  # ITEM_MAP.append(create_item(id=31, ls_item="TestLM", frame=TestLM, actionlist=[ActionManipulator.PICK, ActionManipulator.PLACE], item_model=create_item_model(inner=Rack.SYSMEX_CS2500), lm_id=5, description="LM Test"))
  # Fills the Vision Config List with Projectrelated Data
  # workspaceid and skillid are highly robominds related so probably will not stay like this in the future
  # sample detection: dx and dy are used to calculate the positions in a rack and given by the offset which will be applied in order to assign the sample to a place in the rack
  # create_vision_config(workspace_id="", skill_id="", item_id=-1, capture_pos=p[0,0,0,0,0,0], dx=0, dy=0, target_origin=p[0,0,0,0,0,0], selector="default", description="default")
  # VISION_CONFIG_MAP.append(create_vision_config(workspace_id="96017791-f581-4e9e-93da-6951695fccc8", skill_id="8885cfe1-6784-4293-bd26-52ebdc67bf95", capture_pos=F10_Cap_CF, target_origin=p[0,0,0,0,0,0], item_id=11, description="LM Detect CF"))
  # VISION_CONFIG_MAP.append(create_vision_config(workspace_id="96017791-f581-4e9e-93da-6951695fccc8", skill_id="8885cfe1-6784-4293-bd26-52ebdc67bf95", capture_pos=F8_Cap_Cobas_LM, target_origin=p[0,0,0,0,0,0], item_id=8, description="LM Detect Cobas Racks"))
  # VISION_CONFIG_MAP.append(create_vision_config(workspace_id="8f0ad01c-dc36-4fdd-b295-0b6b4a38b89a", skill_id="afdc9e13-ea83-40d6-a805-bb041453d2e5", capture_pos=F3_Cap_Input, target_origin=F2_uLM_Input, item_id=3, description="Lab Solution Input Capture"))
  # VISION_CONFIG_MAP.append(create_vision_config(workspace_id="96017791-f581-4e9e-93da-6951695fccc8", skill_id="8885cfe1-6784-4293-bd26-52ebdc67bf95", capture_pos=F19_XN550_Cap, target_origin=F18_XN550_Input, item_id=18, description="Input XN550"))
  # VISION_CONFIG_MAP.append(create_vision_config(workspace_id="96017791-f581-4e9e-93da-6951695fccc8", skill_id="8885cfe1-6784-4293-bd26-52ebdc67bf95", capture_pos=F19_XN550_Cap, target_origin=POS_Z, item_id=19, description="LM Detect XN550F"))
  # VISION_CONFIG_MAP.append(create_vision_config(workspace_id="96017791-f581-4e9e-93da-6951695fccc8", skill_id="8885cfe1-6784-4293-bd26-52ebdc67bf95", capture_pos=F10_Cap_CF, target_origin=POS_Z, item_id=10, description="LM Detect CF"))
  # VISION_CONFIG_MAP.append(create_vision_config(workspace_id="96017791-f581-4e9e-93da-6951695fccc8", skill_id="8885cfe1-6784-4293-bd26-52ebdc67bf95", capture_pos=F19_XN550_Cap, target_origin=F20_XN550_Draw, item_id=20, description="Drawer XN550"))
  # VISION_CONFIG_MAP.append(create_vision_config(workspace_id="96017791-f581-4e9e-93da-6951695fccc8", skill_id="8885cfe1-6784-4293-bd26-52ebdc67bf95", capture_pos=F19_XN550_Cap, target_origin=F21_XN550_Btn, item_id=21, description="Button XN550"))
  # VISION_CONFIG_MAP.append(create_vision_config(workspace_id="96017791-f581-4e9e-93da-6951695fccc8", skill_id="8885cfe1-6784-4293-bd26-52ebdc67bf95", capture_pos=TestLMCap, target_origin=p[0,0,0,0,0,0], item_id=30, description="Button XN550"))
  # VISION_CONFIG_MAP.append(create_vision_config(workspace_id="96017791-f581-4e9e-93da-6951695fccc8", skill_id="8885cfe1-6784-4293-bd26-52ebdc67bf95", capture_pos=TestLMCap, target_origin=TestLM, item_id=31, description="Button XN550"))

  # VISION_CONFIG_MAP.append(create_vision_config(workspace_id="96017791-f581-4e9e-93da-6951695fccc8", skill_id="8885cfe1-6784-4293-bd26-52ebdc67bf95", target_origin=p[0,0,0,0,0,0], item_id=11, description="LM Detect CF"))
  # VISION_CONFIG_MAP.append(create_vision_config(workspace_id="96017791-f581-4e9e-93da-6951695fccc8", skill_id="8885cfe1-6784-4293-bd26-52ebdc67bf95", target_origin=p[0,0,0,0,0,0], item_id=8, description="LM Detect Cobas Racks"))
  # VISION_CONFIG_MAP.append(create_vision_config(workspace_id="8f0ad01c-dc36-4fdd-b295-0b6b4a38b89a", skill_id="afdc9e13-ea83-40d6-a805-bb041453d2e5", target_origin=F2_uLM_Input, item_id=3, description="Lab Solution Input Capture"))
  # VISION_CONFIG_MAP.append(create_vision_config(workspace_id="96017791-f581-4e9e-93da-6951695fccc8", skill_id="8885cfe1-6784-4293-bd26-52ebdc67bf95", target_origin=F18_XN550_Input, item_id=18, description="Input XN550"))
  # VISION_CONFIG_MAP.append(create_vision_config(workspace_id="96017791-f581-4e9e-93da-6951695fccc8", skill_id="8885cfe1-6784-4293-bd26-52ebdc67bf95", target_origin=POS_Z, item_id=19, description="LM Detect XN550F"))
  # VISION_CONFIG_MAP.append(create_vision_config(workspace_id="96017791-f581-4e9e-93da-6951695fccc8", skill_id="8885cfe1-6784-4293-bd26-52ebdc67bf95", target_origin=POS_Z, item_id=10, description="LM Detect CF"))
  # VISION_CONFIG_MAP.append(create_vision_config(workspace_id="96017791-f581-4e9e-93da-6951695fccc8", skill_id="8885cfe1-6784-4293-bd26-52ebdc67bf95", target_origin=F20_XN550_Draw, item_id=20, description="Drawer XN550"))
  # VISION_CONFIG_MAP.append(create_vision_config(workspace_id="96017791-f581-4e9e-93da-6951695fccc8", skill_id="8885cfe1-6784-4293-bd26-52ebdc67bf95", target_origin=F21_XN550_Btn, item_id=21, description="Button XN550"))
  # VISION_CONFIG_MAP.append(create_vision_config(workspace_id="96017791-f581-4e9e-93da-6951695fccc8", skill_id="8885cfe1-6784-4293-bd26-52ebdc67bf95", target_origin=p[0,0,0,0,0,0], item_id=30, description="Button XN550"))
  # VISION_CONFIG_MAP.append(create_vision_config(workspace_id="96017791-f581-4e9e-93da-6951695fccc8", skill_id="8885cfe1-6784-4293-bd26-52ebdc67bf95", target_origin=TestLM, item_id=31, description="Button XN550"))

  # local inputrack = find_pattern_by_name("INPUT")
  # INSPECT_CONFIG_MAP.append(create_inspect_config(item_id=3, dx=inputrack.pattern_width[0]/(inputrack.pattern_size[0]-1), dy=inputrack.pattern_width[1]/(inputrack.pattern_size[1]-1), rack_size=inputrack.pattern_size , description="Input Capture"))
  # # Fills the Landmark List with Projectrelated Data
  # # create_landmark(lm_id=0, marker_id=-1, marker_size=0.1, marker_type="aruco_7x7", capture_pos=p[0,0,0,0,0,0], init_frame=p[0,0,0,0,0,0], search_offset=[0,0,0], actual_frame=p[0,0,0,0,0,0], description="")
  # LANDMARK_MAP.append(create_landmark(lm_id=1, marker_id=3, marker_size=0.1, marker_type="aruco_7x7", capture_pos = F10_Cap_CF, init_frame=p[-0.617789, -0.065471, 0.07918, 0.020983, -0.012695, 1.512066], search_offset=[0.15, 0.15, 0.1], actual_frame=p[-0.617789, -0.065471, 0.07918, 0.020983, -0.012695, 1.512066], description="LM CF Lid"))
  # LANDMARK_MAP.append(create_landmark(lm_id=2, marker_id=-1, marker_size=0.0085, marker_type="aruco_4x4", capture_pos = F8_Cap_Cobas_LM, init_frame=p[0,0,0,0,0,0], search_offset=[0.15, 0.15, 0.1], actual_frame=POS_Z, description="LM Cobas Rack Detection"))
  # LANDMARK_MAP.append(create_landmark(lm_id=3, marker_id=0, marker_size=0.1, marker_type="aruco_7x7", capture_pos = F17_Cobas_Cap, init_frame=p[-0.667,-0.194,0.100,0,0,0], search_offset=[0.15, 0.15, 0.1], actual_frame=POS_Z, description="LM Cobas Cap"))
  # LANDMARK_MAP.append(create_landmark(lm_id=4, marker_id=4, marker_size=0.1, marker_type="aruco_7x7", capture_pos = F19_XN550_Cap, init_frame=p[0.124,-0.976,0.355,-0.008,0.025,3.131], search_offset=[0.15, 0.15, 0.1], actual_frame=p[0,0,0,0,0,0], description="LM XN550 Cap"))
  # LANDMARK_MAP.append(create_landmark(lm_id=5, marker_id=0, marker_size=0.1, marker_type="aruco_7x7", capture_pos = TestLMCap, init_frame=p[-0.49,-0.144,0.092,0,-0.008,0.001], search_offset=[0.15, 0.15, 0.1], actual_frame=POS_Z, description="LM Test"))
  # # Configuration of all movement related parameters
  # # create_movement(id=0, hh_approach=POS_Z, h_approach=POS_Z, approach=POS_Z, h_target=POS_Z, target=POS_Z, retract=POS_Z, h_retract=POS_Z, hh_retract=POS_Z, h_frame=POS_Z, frame=POS_Z, speed=1, acceleration=1, description="default")
  # MOVEMENT_MAP.append(create_movement(description="TestLMCap", frame=TestLMCap, actionlist=[ActionManipulator.MOVE_TO]))
  # MOVEMENT_MAP.append(create_movement(description="TestLM", frame=TestLM, actionlist=[ActionManipulator.PICK,ActionManipulator.PLACE],
  #         approach=p[0,0,0.1,0,0,0],
  #         retract=p[0,0,0.1,0,0,0]))
  # MOVEMENT_MAP.append(create_movement(description="Home - MOVE_TO", frame=F1_uLM_Home, actionlist=[ActionManipulator.MOVE_TO]))
  # MOVEMENT_MAP.append(create_movement(description="Input - PICK&PLACE", frame=F2_uLM_Input, actionlist=[ActionManipulator.PICK,ActionManipulator.PLACE],
  #         approach=p[0,0,0.1,0,0,0],
  #         retract=p[0,0,0.1,0,0,0]))
  # MOVEMENT_MAP.append(create_movement(description="Capture Input - MOVE_TO", frame=F3_Cap_Input, actionlist=[ActionManipulator.MOVE_TO]))
  # MOVEMENT_MAP.append(create_movement(description="BIN - PLACE", frame=F4_uLM_Bin, actionlist=[ActionManipulator.PLACE],
  #         approach=p[0,0,0.1,0,0,0],
  #         retract=p[0,0,0.1,0,0,0]))
  # MOVEMENT_MAP.append(create_movement(description="Gripper - Move To", frame=F5_uLM_Gripper, actionlist=[ActionManipulator.MOVE_TO],
  #         approach=p[0,0,0.1,0,0,0]))
  # MOVEMENT_MAP.append(create_movement(description="Gripper - Pick", frame=F5_uLM_Gripper, actionlist=[ActionManipulator.PICK],
  #         retract=p[0,0,0.1,0,0,0]))
  # MOVEMENT_MAP.append(create_movement(description="Gripper - Place", frame=F5_uLM_Gripper, actionlist=[ActionManipulator.PLACE],
  #         approach=p[0,0,0.1,0,0,0]))
  # MOVEMENT_MAP.append(create_movement(description="CobasRack Pick & Place", frame=F6_uLM_Cobas_R, actionlist=[ActionManipulator.PICK,ActionManipulator.PLACE],
  #         approach=p[0,0,0.1,0,0,0],
  #         target=p[0,0,0,0,0,d2r(90)],
  #         retract=p[0,0,0.1,0,0,0]))
  # MOVEMENT_MAP.append(create_movement(description="CobasMagazine Pick & Place", frame=F7_uLM_Coba_Mag, actionlist=[ActionManipulator.PICK,ActionManipulator.PLACE],
  #         approach=p[0,0,0.1,0,0,0],
  #         target=p[0,0,0,0,0,-d2r(90)],
  #         retract=p[0,0,0.1,0,0,0]))
  # MOVEMENT_MAP.append(create_movement(description="Capture Position Cobas Landmarks", frame=F8_Cap_Cobas_LM, actionlist=[ActionManipulator.MOVE_TO]))
  # MOVEMENT_MAP.append(create_movement(description="TaraMagazine - PICK & PLACE", frame=F9_uLM_Tara, actionlist=[ActionManipulator.PICK,ActionManipulator.PLACE],
  #         approach=p[0,0,0.13,0,0,0],
  #         target=p[0,0,0,0,0,-d2r(90)],
  #         retract=p[0,0,0.13,0,0,0]))
  # MOVEMENT_MAP.append(create_movement(description="Capture Position - Centrifuge LM", frame=F10_Cap_CF,actionlist=[ActionManipulator.MOVE_TO]))
  # MOVEMENT_MAP.append(create_movement(description="Pick and Place Racks - Centrifuge Lid", frame=F11_CF_PiPl, actionlist=[ActionManipulator.PICK,ActionManipulator.PLACE],
  #         approach=p[0,0,0.3,0,0,0],
  #         retract=p[0,0,0.3,0,0,0]))
  # MOVEMENT_MAP.append(create_movement(description="Pick and Place Samples - Centrifuge on uLM", frame=F12_uLM_CF_Mag, actionlist=[ActionManipulator.PICK,ActionManipulator.PLACE],
  #         approach=p[0,0,0.13,0,0,0],
  #         retract=p[0,0,0.13,0,0,0]
  #         ))
  # MOVEMENT_MAP.append(create_movement(description="Pick and Place Racks - Centrifuge on uLM", frame=F13_uLM_CF_R, actionlist=[ActionManipulator.PICK,ActionManipulator.PLACE],
  #         approach=p[0,0,0.15,0,0,0],
  #         retract=p[0,0,0.15,0,0,0]
  #         ))

  # MOVEMENT_MAP.append(create_movement(description="Pick and Place Samples XN550 Racks in Device", frame=F18_XN550_Input, actionlist=[ActionManipulator.PICK,ActionManipulator.PLACE],
  #         approach=p[0,0,0.1,0,0,0],
  #         target = p[0,0,0,0,0,d2r(90)],
  #         retract=p[0,0,0.1,0,0,0]
  #         ))
  # MOVEMENT_MAP.append(create_movement(description="Capture LM XN550", frame=F19_XN550_Cap, actionlist=[ActionManipulator.MOVE_TO]))
  # MOVEMENT_MAP.append(create_movement(description="Open XN550 Drawer ", frame=F20_XN550_Draw, actionlist=[ActionManipulator.DRAWER_OPEN],
  #         h_approach=p[0.07,0,0.1,0,0,0],
  #         approach=p[0,0,0.1,0,0,0],
  #         target = p[0,0,0,0,0,d2r(90)],
  #         retract=p[0.07,0,0,0,0,0],
  #         h_retract=p[0.07,0,0.1,0,0,0]
  #         ))
  # MOVEMENT_MAP.append(create_movement(description="Close XN550 Drawer ", frame=F20_XN550_Draw, actionlist=[ActionManipulator.DRAWER_CLOSE],
  #         h_approach=p[0.07,0,0.1,0,0,0],
  #         approach=p[0.07,0,0,0,0,0],
  #         target = p[0,0,0,0,0,d2r(90)],
  #         retract=p[0,0,0.1,0,0,0],
  #         h_retract=p[0.07,0,0.1,0,0,0]
  #         ))
  # MOVEMENT_MAP.append(create_movement(description="Push XN550 Button ", frame=F21_XN550_Btn, actionlist=[ActionManipulator.PUSH],
  #         approach=p[0,0,0.15,0,0,0],
  #         retract=p[0,0,0.15,0,0,0]
  #         ))
  # MOVEMENT_MAP.append(create_movement(description="Capture Position 2 Input", frame=F_Cap_Input2,actionlist=[ActionManipulator.MOVE_TO]))



  $ 19 "Script: SCRIPT Objects V0.1.script"
  #*****************************************************
  # customer          :   INTERNAL
  # project name      :
  #****************************************************
  # controller        :   UR
  # software          :   5.17.3
  #****************************************************
  # author            :   P. Koehnke
  # Copyright (c)     :   United Robotics Group
  #                       An der Riede 2
  #                       28816 Stuhr
  #                       Germany
  #****************************************************
  # description       :   object database
  # version:      	:   0.1
  # created           :   09.10.2024
  # updated           :
  #****************************************************
  # modifications     :
  #
  # date              :
  # name              :
  # reason            :
  #****************************************************

  def create_object_2(id=0, name="", type=0, dimension=struct(length=0, width=0, height=0, diameter=0), gripper_offset=p[0,0,0,0,0,0]):
      return struct(id=id, name=name, type=type, dimension=dimension, gripper_offset=gripper_offset)
  end

  OBJ = create_object_2()
  OBJs = make_list(0, create_object_2(), 50)

  OBJs.append(create_object_2(id=1, name="rack centrifuge", type=1, dimension=struct(length=0, width=0, height=0.106, diameter=0.020), gripper_offset=p[0,0,0.095,0,0,2.356]))
  OBJs.append(create_object_2(id=2, name="sample tube 1", type=2, dimension=struct(length=0, width=0, height=0.106, diameter=0.015), gripper_offset=p[0,0,0,0,0,0]))
  OBJs.append(create_object_2(id=3, name="rack sarstedt", type=3, dimension=struct(length=0, width=0, height=0.100, diameter=0.020), gripper_offset=p[0,0,0,0,0,0]))
  OBJs.append(create_object_2(id=4, name="Lab bottle", type=4, dimension=struct(length=0, width=0, height=0.100, diameter=0.030), gripper_offset=p[0,0,0.2,0,0,0]))
  OBJs.append(create_object_2(id=5, name="Vial", type=5, dimension=struct(length=0, width=0, height=0.100, diameter=0.0275), gripper_offset=p[0,0,0,0,0,0]))
  OBJs.append(create_object_2(id=6, name="Container", type=6, dimension=struct(length=0.0, width=0.0, height=0, diameter=0.0), gripper_offset=p[0,0,0,0,0,0]))
  OBJs.append(create_object_2(id=7, name="Target_container", type=7, dimension=struct(length=0.06, width=0.06, height=0.134, diameter=0.05), gripper_offset=p[0,0,0,0,0,0]))
  OBJs.append(create_object_2(id=8, name="Spatula", type=8, dimension=struct(length=0.03, width=0.03, height=0.23, diameter=0.05), gripper_offset=p[0,0,0,0,0,0]))
  OBJs.append(create_object_2(id=9, name="rack pipet", type=9, dimension=struct(length=0.03, width=0.03, height=0.23, diameter=0.05), gripper_offset=p[0,0,0,0,0,0]))

  def create_jig_2(id=0, name="", type=0, capacity=0, jig_offset=p[0,0,0,0,0,0]):
      # iformation about used jigs
      return struct(id=id, name=name, type=type, capacity=capacity, jig_offset=jig_offset)
  end

  JIG2 = create_jig_2()
  JIGs = make_list(0, create_jig_2(), 20)

  JIGs.append(create_jig_2(id=1, name="3FG", type=1, capacity=1, jig_offset=p[0,0,0,0,0,0]))
  JIGs.append(create_jig_2(id=2, name="jig input", type=2, capacity=1, jig_offset=p[0,0,0,0,0,-3.927]))
  JIGs.append(create_jig_2(id=3, name="jig output", type=3, capacity=1, jig_offset=p[0,0,0,0,0,0.78]))
  JIGs.append(create_jig_2(id=6, name="jig bin", type=6, capacity=1, jig_offset=p[0,0,0,0,0,0]))
  JIGs.append(create_jig_2(id=7, name="jig sarstedt racks", type=7, capacity=1, jig_offset=p[0,0,-0.02,0,0,0]))
  JIGs.append(create_jig_2(id=8, name="NoK Bin", type=8, capacity=1, jig_offset=p[0,0,0,0,0,0]))
  JIGs.append(create_jig_2(id=9, name="Pick bott jig", type=9, capacity=1, jig_offset=p[0,0,0,0,0,0]))
  JIGs.append(create_jig_2(id=10, name="Place bott jig", type=10, capacity=1, jig_offset=p[0,0,0,0,0,0]))
  JIGs.append(create_jig_2(id=11, name="bottle shake jig", type=11, capacity=1, jig_offset=p[0,0,0,0,0,0]))
  JIGs.append(create_jig_2(id=12, name="Pick Vial jig", type=12, capacity=1, jig_offset=p[0,0,0,0,0,0]))
  JIGs.append(create_jig_2(id=13, name="Place Vial jig", type=13, capacity=1, jig_offset=p[0,0,0,0,0,0]))
  JIGs.append(create_jig_2(id=14, name="Liquid transfer jig", type=14, capacity=1, jig_offset=p[0,0,0,0,0,0]))
  JIGs.append(create_jig_2(id=15, name="Pick station jig", type=15, capacity=1, jig_offset=p[0,0,0,0,0,0]))
  JIGs.append(create_jig_2(id=16, name="Place station jig", type=16, capacity=1, jig_offset=p[0,0,0,0,0,0]))
  JIGs.append(create_jig_2(id=17, name="Weigh station jig", type=17, capacity=1, jig_offset=p[0,0,0,0,0,0]))
  JIGs.append(create_jig_2(id=18, name="Pick station 1", type=18, capacity=1, jig_offset=p[0,0,0,0,0,0]))
  JIGs.append(create_jig_2(id=19, name="Pick station 2", type=19, capacity=1, jig_offset=p[0,0,0,0,0,0]))
  JIGs.append(create_jig_2(id=20, name="Pick station 3", type=20, capacity=1, jig_offset=p[0,0,0,0,0,0]))
  JIGs.append(create_jig_2(id=21, name="Tilt station jig", type=21, capacity=1, jig_offset=p[0,0,0,0,0,0]))
  $ 26 "Script: Powder_all.script"
  global SERVER_IP   = "192.168.12.139"
  global SERVER_PORT = 3002

  global POTS_IP   = "192.168.12.111"
  global POTS_PORT = 80

  global container_id = 0
  global powder_id  = 0
  global bulk_density = 0
  global H          = 0
  global H_c          = 0
  global mouth_d     = 0
  global mouth_sh    = 0
  global length_c     = 0
  global diameter   = 0
  global empty_weight_g  = 0
  global volume_ml    = 0
  global shape_code   = 0
  global flow_code   = 0
  global shape = ""
  global Flowability = ""
  global full_weight_g = 0
  global cent_edge = 0
  global pick_2_base = 0.2 # distance from tcp to base of picking table
  global wall_thickness = 0.005

  def read_db_data():

    socket_open(SERVER_IP, SERVER_PORT)
    sleep(0.5)
    socket_send_string("GET_DATACODE_FLOATS")
    sleep(5)

    local fl = socket_read_ascii_float(14)
    socket_close()

    global container_id = fl[1]
    global powder_id = fl[2]
    global bulk_density = fl[3]
    global H          = fl[4]/1000
    global H_c          = fl[5]/1000
    global mouth_d     = fl[6]/1000
    global mouth_sh    = fl[7]/1000
    global length_c     = fl[8]/1000
    global diameter   = fl[9]/1000
    global empty_weight_g = fl[10]
    global volume_ml    = fl[11]
    global full_weight_g = fl[12]
    global flow_code   = fl[13]
    global shape_code   = fl[14]

  	if (flow_code == 1.0):
  	  global Flowability = "MEDIUM"
  	elif (flow_code == 2.0):
  	  global Flowability = "LOW"
  	else:
  	  global Flowability = "HIGH"
  	end

    if ( shape_code == 1.0):
  	shape = "cylindrical"
  	cent_edge =  diameter
    else:
  	shape = "cubical"
  	cent_edge =  length_c
    end

  end

  def send_picking_info(Pow_name, target_weight):
    socket_open(SERVER_IP, SERVER_PORT)
    cmd = "PICK:"+Pow_name+";"+to_str(target_weight)
    socket_send_string(cmd)
    sleep(0.1)
    socket_close()
  end

  #### POTS ####
  def tilt_send(angle):
  	socket_open(POTS_IP, POTS_PORT)
  	angle = 92.0 - angle
  	socket_send_string("Tilt,"+to_str(angle)+",0")
  	sync()
  	sleep(0.5)
  	socket_close()
  end

  def Motors_off():
  	socket_open(POTS_IP, POTS_PORT)
  	socket_send_string("Off,0,0")
  	sync()
  	sleep(0.5)
  	socket_close()
  end

  def Rotate():
  	socket_open(POTS_IP, POTS_PORT)
  	socket_send_string("FullRotation, 1, 2000")
  	sync()
  	sleep(0.5)
  	socket_close()
  end

  def CCW_Rotate():
  	socket_open(POTS_IP, POTS_PORT)
  	socket_send_string("FullRotation, -1, 2000")
  	sync()
  	sleep(0.5)
  	socket_close()
  end

  def tilt_to_home():
  	socket_open(POTS_IP, POTS_PORT)
  	socket_send_string("Home,0,0")
  	sync()
  	sleep(0.5)
  	socket_close()
  end
  #######
  def vibration_1():
  	set_analog_out(0,0.4)
  	sleep(1)
  	set_analog_out(0,0.0)
  	sleep(0)
  end

  def vibration_2():
  	set_analog_out(0,0.8)
  	sleep(0.8)
  	set_analog_out(0,0.0)
  	sleep(0.2)
  end

  def vibration_3():
  	set_analog_out(0,0.4)
  	sleep(0.5)
  	set_analog_out(0,0.0)
  	sleep(0.3)
  end

  def vibration_4():
  	set_analog_out(0,0.4)
  	sleep(0.6)
  	set_analog_out(0, 0.0)
  	sleep(0.5)
  end

  ##################

  global gear_2_holder = 0.018
  global gain_per_percent = 0.5
  global w_dosed_total = 0.0
  global last_scale = 0.0
  global tilt_angle_sent = 0.0
  global level = 0.0
  global target_g = 0.0
  global angle_max = 60
  global angle_min = 10
  global hinge_2_base = 0.0421
  global TCP_2_tip_x = 0.0047
  global spatula_len = 0.182
  global spatula_offset = p[TCP_2_tip_x,0,spatula_len,0,0,0]
  global SPATULA_L_VOL_ML = 5.0        # 1 teaspoon = 5 mL
  global SPATULA_M_VOL_ML = 1.25       # 1/4 teaspoon = 1.25 mL
  global SPATULA_S_VOL_ML = 0.15625    # 1/32 teaspoon = 0.15625 mL
  global SPATULA_FLAT_M_VOL_ML  = 2.2
  global SPATULA_FLAT_S_VOL_ML  = 1.2   #based on caluclations using rho = m/V
  global ry_deg_safe = 0
  global ry_deg = 0



  def clamp(x, lo, hi):
  	if(x<lo):
  		return lo
  	elif (x>hi):
  		return hi
  	else:
  		return x
  	end
  end

  def compute_level_percent(W_now, weight_value):   # W_now = container+powder, weight_value = live scale reading
      local delta = weight_value - last_scale

      if (delta < 0.0):
          delta = 0.0
      end

      global w_dosed_total = w_dosed_total + delta
      global last_scale = weight_value     # update the last scale reading

      local W_eff = W_now - w_dosed_total
      if (W_eff <  empty_weight_g):
          W_eff =  empty_weight_g
      end

      # Compute powder level %
      level = 100.0 * (W_eff -  empty_weight_g) / (full_weight_g -  empty_weight_g)

      # Clamp to 0–100
      level = clamp(level, 0, 100)
    textmsg("deb 1 = ", level)
      return level
  end

  def deg2rad(d):
  	return d*3.141592/180
  end

  def my_abs(val):
  	if (val<0):
  		return -val
  	else:
  		return val
  	end
  end

  def compute_tilt_deg(level_percent):
  	angle = angle_min + gain_per_percent*(100.0-level_percent)

    	textmsg("deb 2 = ", angle)
  	return clamp(angle, angle_min, angle_max)
  end

  def tilt(level_percentage):
  	new_angle = compute_tilt_deg(level_percentage)
  	global angle_rel = new_angle - tilt_angle_sent

  	if my_abs(angle_rel)>2.0:
  		tilt_send(new_angle)
  		global angle_deg = new_angle
  		global tilt_angle_sent = new_angle
  		global p_center_vertical = center_pose()
  		global p_center = updated_center_pose(p_center_vertical, angle_deg)
  	end

  	if (level_percentage<85.0):
  		tilt_send(angle_deg)
  	end
  end

  def compute_scoop_depth(level):
    return ((100.0-level)/100.0)*(H -mouth_sh )
  end

  def map_tilt_to_ry_deg(container_deg, level):

  	if (Flowability == "HIGH" or Flowability == "MEDIUM"):
  		global scoop_depth = compute_scoop_depth(level)
  		safe_scoop_pivot = (mouth_d  - spatula_depth)/(scoop_depth+mouth_sh+spatula_mid)
  		global ry_deg_safe = asin(safe_scoop_pivot)
  		global ry_deg = 90-container_deg
  	else:
  		global scoop_depth = compute_scoop_depth(level)
  		safe_scoop_pivot = (mouth_d  - spatula_depth)/(scoop_depth+mouth_sh+spatula_mid )
  		global ry_deg_safe = asin(safe_scoop_pivot)
  		global ry_deg = 90-container_deg
  	end
  	return [ry_deg_safe,ry_deg]
  end

  def get_scoop_weight(spatula, bulk_density):

  	local vol = 0

  	if (spatula == "spatula_L"):
  		vol = SPATULA_L_VOL_ML
  		global spatula_depth = 0.015
  		global spatula_mid   = 0.016
  		global spatula_ry    = 0.0

  	elif (spatula == "spatula_M"):
  		vol = SPATULA_M_VOL_ML
  		global spatula_depth = 0.010
  		global spatula_mid   = 0.0105
  		global spatula_ry    = 0.0

  	elif (spatula == "spatula_S"):
  		vol = SPATULA_S_VOL_ML
  		global spatula_depth = 0.008
  		global spatula_mid   = 0.0063
  		global spatula_ry    = 0.0

  	elif (spatula == "spatula_flat_M"):
  		vol = SPATULA_FLAT_M_VOL_ML
  		global spatula_depth = 0.001
  		global spatula_mid   = 0.002
  		global spatula_ry    = 10.0

  	elif (spatula == "spatula_flat_S"):
  		vol = SPATULA_FLAT_S_VOL_ML
  		global spatula_depth = 0.005
  		global spatula_mid   = 0.016
  		global spatula_ry    = 2.0

  	else:
  		textmsg("Unknown spatula type")
  		return 0.0
  	end
  	global target_g = vol * bulk_density
  	return target_g

  end

  def select_spatula(Flowability, level, diff, bulk_density, mouth_d ):

      local k = 1.1

      global powder_height = (H  - mouth_sh ) * level/100

      if (Flowability == "LOW"):

          local gFM = get_scoop_weight("spatula_flat_M", bulk_density)

          local level_ok_FM = (spatula_mid  < powder_height)
          local diff_ok_FM  = (diff > k * gFM)

          local flatM_ok = level_ok_FM and diff_ok_FM

          if (flatM_ok):
              return "spatula_flat_M"
          else:
              return "spatula_flat_S"
          end

      end

      local gL = get_scoop_weight("spatula_L", bulk_density)

      local mouth_ok_L = (mouth_d  >= 0.05)
      local level_ok_L = (spatula_mid < powder_height)
      local diff_ok_L  = (diff > k * gL)

      local large_ok = mouth_ok_L and level_ok_L and diff_ok_L

      local gM = get_scoop_weight("spatula_M", bulk_density)

      local level_ok_M = (spatula_mid < powder_height)
      local diff_ok_M  = (diff > k * gM)

      local medium_ok = level_ok_M and diff_ok_M

      if (large_ok):
          return "spatula_L"

      elif (medium_ok):
          return "spatula_M"

      else:
          return "spatula_S"
      end

  end

  def after_scoop():

  	set_analog_out(0,0.0)
  	tilt_send(angle_deg)
  	sleep(0.5)
  	movel(lifted_pose, a=0.05, v=0.2)
  	movel(tilted_pose_in_base2, a=0.05, v=0.2)
  	set_analog_out(0,0.4)
  	movel(pose_trans(tilted_pose_in_base2, p[0,0,0,0,0,2.0]), a=0.05, v=0.2)
  	set_analog_out(0,0.0)
  	movel(tilted_pose_in_base2, a=0.05, v=0.2)
  	movel(lifted_pose, a=0.05, v=0.2)
  	tilt_to_home()
  end

  def center_pose():
  	global p_translated = container_place
  	#global p_translated = pots_axis_temp

  	#cx = p_translated[0]
  	#cy = p_translated[1]
  	#cz = p_translated[2]

  	global p_center_vertical_temp = pose_trans(p_translated, p[0,0,0, deg2rad(90), 0, 0])
  	cx = p_center_vertical_temp[0]
  	cy = p_center_vertical_temp[1]
  	cz = p_center_vertical_temp[2]
  	rx = p_center_vertical_temp[3]
  	ry = p_center_vertical_temp[4]
  	rz = p_center_vertical_temp[5]

  	global p_center_vertical_temp = p[cx,cy,cz, 0, 0, rz]
  	trans_rel = p[0,0,-pick_2_base+H,0,0,0]
  	global p_center_vertical =  pose_trans(p_center_vertical_temp, trans_rel)
  	return p_center_vertical
  end

  def updated_center_pose(p_center_vertical, angle_deg):
  	hinge_pose = pose_trans(p_center_vertical, p[0,0,-hinge_2_base-gear_2_holder-H ,0,0,0])
  	local_rel = pose_trans(pose_inv(hinge_pose), p_center_vertical)

  	rot_tilt = p[0,0,0, -deg2rad(angle_deg),0,0]
  	local_rel_tilted = pose_trans(rot_tilt, local_rel)

  	global p_center = pose_trans(hinge_pose, local_rel_tilted)
  	return p_center
  end

  def scoop_powder(p_center):
  	vibration_voltage = 0.4
  	global scoop_radius_default = 0.0


  	scoop_radius_default = mouth_d /2 - spatula_depth
  	scoop_safe_entry_pose = pose_trans(p_center, p[-TCP_2_tip_x,0,spatula_len+0.05,0,0,0])
  	scoop_entry_pose = pose_trans(p_center, p[-TCP_2_tip_x,0,spatula_len,0,0,0])

  	movel(scoop_safe_entry_pose, a=0.1, v=0.25)
  	movel(scoop_entry_pose, a=0.1, v=0.25)

  	scoop_start_rel_int = p[0, 0, -mouth_sh , 0, 0, 0]
  	scoop_start_pose_int = pose_trans(scoop_entry_pose, scoop_start_rel_int)

  	movel(scoop_start_pose_int, a=0.1, v=0.25)

  	#local ry_deg = map_tilt_to_ry_deg(angle_deg,level)
  	local ry_result = map_tilt_to_ry_deg(angle_deg,level)
  	global ry_safe = ry_result[0]
  	global ry = deg2rad(ry_result[1])

  	if (spatula_mid < powder_height):

  		global total_depth = mouth_sh + scoop_depth + spatula_mid
  		global total_depth = clamp(total_depth, 0, H - spatula_mid)
  		scoop_start_rel = p[scoop_radius_default, 0, -total_depth, 0, 0, 0]

  		rot_mid = p[0, 0, 0, 0, 0, 0.785]
  		rot_end = p[0, 0, 0, 0, 0, 1.5708]

  		scoop_via_rel = pose_trans(rot_mid, scoop_start_rel)
  		scoop_end_rel = pose_trans(rot_end, scoop_start_rel)

  		scoop_start_pose = pose_trans(scoop_entry_pose, scoop_start_rel)
  		scoop_via_pose = pose_trans(scoop_entry_pose, scoop_via_rel)
  		scoop_end_pose = pose_trans(scoop_entry_pose, scoop_end_rel)

  		movel(scoop_start_pose, a=0.5, v=0.3)

  		if (level<90.0):
  			Rotate()
  		end

  		movec(scoop_via_pose, scoop_end_pose, a=0.03, v=0.02)
  		sleep(1.0)


  		# safe_retention
  		local pivot_pose = pose_trans(scoop_end_pose, p[0,0,total_depth-spatula_len,0,0,0])
  		local end_rel = pose_trans(pose_inv(pivot_pose), scoop_end_pose)
  		local end_rel_tilted = pose_trans(end_rel, p[0, 0, 0, 0, ry_safe, 0])
  		global tilted_pose_in_base = pose_trans(pivot_pose, p[0,0,0,end_rel_tilted[3],end_rel_tilted[4], end_rel_tilted[5]])
  		global tilted_pose_in_base = pose_trans(tilted_pose_in_base, p[0, 0, spatula_len-total_depth, 0, 0, 0])
  		# sptula pivoted around the container rim of the mouth at ry_safe
  		movel(tilted_pose_in_base, a=0.03, v=0.1)

  		global safe_x = sin(ry_safe)*(scoop_depth - (mouth_d -spatula_depth)/tan(90-ry_safe/2))
  		global safe_z = cos(ry_safe)*(scoop_depth - (mouth_d -spatula_depth)/tan(90-ry_safe/2))

  		local safe_up = pose_trans(tilted_pose_in_base, p[-safe_x,0,safe_z,0,0,0])
  		movel(safe_up, a=0.03, v=0.1)

  		# full exit
  		local pivot_pose2 = pose_trans(tilted_pose_in_base, p[0,0,total_depth-spatula_len,0,0,0])
  		local end_rel2 = pose_trans(pose_inv(pivot_pose2), tilted_pose_in_base)
  		#popup("is the spatula crashing front? ", blocking = True)
  		local end_rel_tilted2 = pose_trans(end_rel2, p[0, 0, 0, 0, ry-ry_safe, 0])
  		global tilted_pose_in_base2 = pose_trans(pivot_pose2, p[0,0,0,end_rel_tilted2[3],end_rel_tilted2[4], end_rel_tilted2[5]])
  		global tilted_pose_in_base2 = pose_trans(tilted_pose_in_base2, p[-TCP_2_tip_x, 0, spatula_len-scoop_radius_default-spatula_mid, 0, 0, 0])
  		# spaula exited at center of the mouth at ry
  		movel(tilted_pose_in_base2, a=0.03, v=0.1)
  		#popup("is the spatula crashing at mouth? ", blocking = True)

  	else : # emptying logic
  		spatula_base = pose_trans(scoop_entry_pose, p[0, 0, -H+wall_thickness, 0, 0, 0])
  		local pivot_pose = pose_trans(scoop_entry_pose, p[0,0,-spatula_len,0,0,0])
  		# tilt inwards
  		global in_angle = atan((cent_edge-2*spatula_depth)/(2*H))
  		spatula_tilt_rel = pose_trans(pose_inv(pivot_pose), spatula_base)

  		spatula_tilt = pose_trans(spatula_tilt_rel, p[0, 0, 0, in_angle, 0, 0])
  		global tilted_pose = pose_trans(pivot_pose, p[0,0,0,spatula_tilt[3],spatula_tilt[4], spatula_tilt[5]])

  		global tilted_pose = pose_trans(tilted_pose, p[0,0,spatula_len-H+wall_thickness,0,0,0])

  		movel(tilted_pose,a=0.1, v=0.25)
  		CCW_Rotate()

  		rotate90=pose_trans(tilted_pose,p[0,0,0,0,0,1.5708])

  		movel(rotate90, a=0.1, v=0.1)
  		#popup("is the spatula crashing front? ", blocking = True)
  		movel(pose_trans(scoop_start_pose_int,p[0,0,0,0,0,1.5708]), a=0.03, v=0.1)
  		# full exit
  		#local pivot_pose2 = pose_trans(scoop_entry_pose, p[0,0,-spatula_len,0,0,0])
  		local end_rel2 = pose_trans(pose_inv(scoop_entry_pose), rotate90)
  		local end_rel_tilted2 = pose_trans(end_rel2, p[0, 0, 0, 0, ry+in_angle, 0])
  		global tilted_pose_in_base2 = pose_trans(pivot_pose, p[0,0,0,end_rel_tilted2[3],end_rel_tilted2[4], end_rel_tilted2[5]])
  		global tilted_pose_in_base2 = pose_trans(tilted_pose_in_base2, p[0, 0, spatula_len, 0, 0, 0])
  		# sptula exited at center of the mouth at ry
  		movel(tilted_pose_in_base2, a=0.03, v=0.1)
  		#popup("is the spatula crashing at mouth? ", blocking = True)
  	end

  	if (spatula=="spatula_flat_S" or spatula=="spatula_S"):
  		vibration_3()
  		local ry_level = deg2rad(20)
  	elif (spatula == "spatula_M"):
  		vibration_3()
  		local ry_level = deg2rad(25)
  	else:
  		vibration_2()
  		local ry_level = deg2rad(15)
  	end

  	# remove excess
  	local pivot_pose_level = pose_trans(tilted_pose_in_base2, p[0,0,-spatula_len,0,0,0])
  	local end_rel_level = pose_trans(pose_inv(pivot_pose_level), tilted_pose_in_base2)
  	#local ry_level = ry/1.5
  	#local ry_level = deg2rad(15)
  	local end_rel_tilted_level = pose_trans(end_rel_level, p[0, 0, 0, 0, -ry_level, 0])
  	local end_rel_tilted_level2 = pose_trans(pivot_pose_level, p[0, 0, 0,end_rel_tilted_level[3],end_rel_tilted_level[4], end_rel_tilted_level[5]])
  	local end_rel_tilted_level2 = pose_trans(end_rel_tilted_level2, p[0,0,spatula_len-spatula_mid,0,0,0])
  	movel(end_rel_tilted_level2, a=0.03, v=0.1)

  	movel(tilted_pose_in_base2, a=0.03, v=0.1)
  	set_analog_out(0, 0.0)
  	#popup("safe out + moving towards beaker", title = "Pause", blocking = True)
  	global lifted_pose = pose_trans(tilted_pose_in_base2, p[-0.04,0,0.04,0,0,0]) # safety distance away from the container

  	movel(lifted_pose, a=0.03, v=0.1)
  	tilt_to_home()
  end

  def auto_tilt_and_scoop(W_now, target_weight, weight_value):
  	global level = compute_level_percent(W_now, weight_value)

  	global spatula = select_spatula(Flowability, level, diff, bulk_density, mouth_d )
  	textmsg("deb 4 8 = ", spatula)
  	global target_g = get_scoop_weight(spatula, bulk_density)

    	#textmsg("deb 4 = ", target_g)
  	#send_scoop_target_info()

  	global scoop_depth = compute_scoop_depth(level)

    	textmsg("deb 5 = ", scoop_depth)
  	#tilt_to_home()
  	#sleep(1.5)
  	tilt(level)
  	#sleep(1.5)
    	#popup("is the pots tilted? ", blocking = True)
    	#textmsg("deb 6 = ", p_center)
  	scoop_powder(p_center)

    	textmsg("deb 7 - sucess")
  end
  $ 27 "Script: Weight_scale_socket_s.script"
  global s_depth = 0
  global s_length =0
  global s_volume = 0
  global ry_theta  = 0

  def get_weight():
  	socket_open(SERVER_IP,SERVER_PORT)
  	sleep(0.2)
  	textmsg("socket opened successfully!")
  	socket_send_string("GET_WEIGHT")
  	sleep(0.2)
  	sync()
  	sleep(0.2)
  	receiveFromServ = socket_read_ascii_float(6)
  	sleep(1)
  	#while (receiveFromServ[0] <1):
  		#receiveFromServ = socket_read_ascii_float(1)
  		#sleep(1)
  		#textmsg("retrying read:", receiveFromServ)
  	#end
  	textmsg("Received weight:", receiveFromServ[1])
  	sleep(0.2)
  	socket_close()
  	sleep(0.2)
  	return receiveFromServ[1]
  end

  def tare_scale():
  	socket_open(SERVER_IP,SERVER_PORT)
  	socket_send_string("TARE")
  	sleep(2)
  	socket_close()
  end

  def zero_scale():
  	socket_open(SERVER_IP,SERVER_PORT)
  	socket_send_string("ZERO")
  	sleep(0.5)
  	socket_close()
  end

  def log_weight():
  	socket_open(SERVER_IP,SERVER_PORT)
  	socket_send_string("LOG_WEIGHT")
  	sleep(0.5)
  	socket_close()
  end

  def send_target_info():
  	socket_open(SERVER_IP,SERVER_PORT)
  	socket_send_string("SET_TARGET:" + to_str(target_weight))
  	sleep(0.2)
  	socket_close()
  end
  def send_powder_info():
  	socket_open(SERVER_IP,SERVER_PORT)
  	socket_send_string("SET_POWDER:" + Pow_name)
  	sleep(0.2)
  	socket_close()
  end
  def send_spatula_info():
  	socket_open(SERVER_IP,SERVER_PORT)
  	socket_send_string("SET_SPATULA:" + spatula)
  	#sleep(1)

  	#local fl = socket_read_ascii_float(4)
    	#socket_close()

    	#global s_depth = fl[1]
    	#global s_length = fl[2]
   	#global s_volume = fl[3]
   	#global ry_theta  = fl[4]
  	sleep(0.2)

  end

  def send_level_info():
  	socket_open(SERVER_IP,SERVER_PORT)
  	socket_send_string("SET_LEVEL:" + to_str(level))
  	sleep(0.2)
  	socket_close()
  end

  def send_weight_info():
    socket_open(SERVER_IP, SERVER_PORT)
    #rq_open_and_wait()
    cmd = "GET_CONT_WEIGHT"
    socket_send_string(cmd)
    sync()
    sleep(0.5)
    receiveFromSer = socket_read_ascii_float(1)
    socket_close()
    return receiveFromSer[1]
  end

  $ 28 "BeforeStarts"
  $ 29 "uLM"
  $ 30 "CMD_Stop≔ False "
  global CMD_Stop=  False
  $ 31 "CMD_Abort≔ False "
  global CMD_Abort=  False
  $ 32 "CMD_Clear≔ False "
  global CMD_Clear=  False
  $ 33 "STATE≔1"
  global STATE=1
  $ 34 "STATE_Info≔''"
  global STATE_Info=""
  $ 35 "ARM_Referenced≔ False "
  global ARM_Referenced=  False
  $ 36 "zero_ftsensor()"
  zero_ftsensor()
  $ 37 "poses init"
  $ 38 "PSE_A≔p[0,0,0,0,0,0]"
  global PSE_A=p[0,0,0,0,0,0]
  $ 39 "PSE_A_H≔p[0,0,0,0,0,0]"
  global PSE_A_H=p[0,0,0,0,0,0]
  $ 40 "PSE_R≔p[0,0,0,0,0,0]"
  global PSE_R=p[0,0,0,0,0,0]
  $ 41 "PSE_R_H≔p[0,0,0,0,0,0]"
  global PSE_R_H=p[0,0,0,0,0,0]
  $ 42 "PSE_T≔p[0,0,0,0,0,0]"
  global PSE_T=p[0,0,0,0,0,0]
  $ 43 "PSE_T_H≔p[0,0,0,0,0,0]"
  global PSE_T_H=p[0,0,0,0,0,0]
  $ 44 "PSE_C_E≔p[0,0,0,0,0,0]"
  global PSE_C_E=p[0,0,0,0,0,0]
  $ 45 "PSE_C_H≔p[0,0,0,0,0,0]"
  global PSE_C_H=p[0,0,0,0,0,0]
  $ 46 "PSE_C_S≔p[0,0,0,0,0,0]"
  global PSE_C_S=p[0,0,0,0,0,0]
  $ 47 "init_home_by_cartesian_pose(p[0,-0.400,0.300,0,0,0])"
  init_home_by_cartesian_pose(p[0,-0.400,0.300,0,0,0])
  $ 48 "Clearing"
  $ 49 "reset_error()"
  reset_error()
  $ 50 "reset_warning()"
  reset_warning()
  $ 51 "uGo"
  $ 53 "ugo_init( True ,'http://192.168.12.120:10001')"
  ugo_init(  True  ,"http://192.168.12.120:10001")
  $ 54 "ugo_update_outputs()"
  ugo_update_outputs()
  $ 55 "App"
  $ 56 "'ADD APPLICATION SPECIFIC COMMANDS'"
  # 'ADD APPLICATION SPECIFIC COMMANDS'
  $ 57 "Tools"
  $ 58 "OBJ_Picked≔gripper_has_object()"
  global OBJ_Picked=gripper_has_object()
  $ 59 "If OBJ_Picked"
  if (OBJ_Picked):
    # begin: URCap Program Node
    #   Source: Robotiq_Grippers, 3.17.0.105337, Robotiq Inc.
    #   Type: Gripper Activate
    $ 60 "Gripper Activate"

    kill rq_gripper_communication_thread
    rq_gripper_communication_thread_started = False
    rq_close_gripper_socket("1")
    rq_close_gripper_socket("2")
    rq_close_gripper_socket("3")
    rq_close_gripper_socket("4")

    rq_init_comm_if_connected(9, "1")
    rq_init_comm_if_connected(2, "2")
    rq_init_comm_if_connected(3, "3")
    rq_init_comm_if_connected(4, "4")
    rq_print_connected_grippers()
    rq_gripper_communication_thread = run rq_gripper_communication()

    while(not rq_gripper_communication_thread_started):
        sleep(0.008)
    end

    rq_set_max_current_for_all_grippers()

    reset_and_activate = False

    rq_activate_all_grippers(False)
    # end: URCap Program Node
  else:
    $ 61 "Else" "noBreak"
    # begin: URCap Program Node
    #   Source: Robotiq_Grippers, 3.17.0.105337, Robotiq Inc.
    #   Type: Gripper Activate
    $ 62 "Gripper Reset and Activate"

    kill rq_gripper_communication_thread
    rq_gripper_communication_thread_started = False
    rq_close_gripper_socket("1")
    rq_close_gripper_socket("2")
    rq_close_gripper_socket("3")
    rq_close_gripper_socket("4")

    rq_init_comm_if_connected(9, "1")
    rq_init_comm_if_connected(2, "2")
    rq_init_comm_if_connected(3, "3")
    rq_init_comm_if_connected(4, "4")
    rq_print_connected_grippers()
    rq_gripper_communication_thread = run rq_gripper_communication()

    while(not rq_gripper_communication_thread_started):
        sleep(0.008)
    end

    rq_set_max_current_for_all_grippers()

    reset_and_activate = True

    rq_activate_all_grippers(True)
    # end: URCap Program Node
  end
  $ 63 "zero_ftsensor()"
  zero_ftsensor()
  $ 64 "EXTT"
  $ 65 "Set GRP_3F_Enable=Off"
  set_standard_digital_out(4, False)
  $ 66 "Set BarcodeTrigger=Off"
  set_standard_digital_out(6, False)
  $ 67 "Set GRP_3F_Decap=Off"
  set_standard_digital_out(3, False)
  $ 68 "Set GRP_3F_Cap=Off"
  set_standard_digital_out(2, False)
  $ 69 "Set GRP_3F_Open=Off"
  set_standard_digital_out(5, False)
  $ 70 "PSE_T≔get_tool_free_pose(dir=[0,0,0.150], move_in_base_frame=True)"
  global PSE_T=get_tool_free_pose(dir=[0,0,0.150], move_in_base_frame=True)
  $ 71 "If is_reachable(Base_const, [PSE_T])"
  if (is_reachable(p[0.0,0.0,0.0,0.0,0.0,0.0], [PSE_T])):
    $ 72 "MoveL"
    $ 73 "PSE_T" "breakAfter"
    movel(PSE_T, a=1.2, v=0.15)
  end
  $ 75 "powder dispensing variable init"
  $ 76 "Start_thread≔ False "
  global Start_thread=  False
  $ 77 "vib_thread≔ False "
  global vib_thread=  False
  $ 78 "w_full_thread≔ False "
  global w_full_thread=  False
  $ 79 "d_cc≔0.07"
  global d_cc=0.07
  $ 80 "kp≔0.0015"
  global kp=0.0015
  $ 81 "ki≔0.0001"
  global ki=0.0001
  $ 82 "kd≔0.01"
  global kd=0.01
  $ 83 "dt≔0.02"
  global dt=0.02
  $ 84 "Integral_error≔0"
  global Integral_error=0
  $ 85 "current_error≔0"
  global current_error=0
  $ 86 "previous_error≔0"
  global previous_error=0
  $ 87 "tilt_increment≔0"
  global tilt_increment=0
  $ 88 "tilt_angle≔0"
  global tilt_angle=0
  $ 89 "diff≔0"
  global diff=0
  $ 95 "tilt_to_home()"
  tilt_to_home()
  $ 96 "switch_spat_M≔ True "
  global switch_spat_M=  True
  $ 97 "switch_spat_S≔ True "
  global switch_spat_S=  True
  $ 98 "switch_spat_F_M≔ True "
  global switch_spat_F_M=  True
  $ 99 "switch_spat_F_S≔ True "
  global switch_spat_F_S=  True
  $ 100 "last_scale≔0"
  global last_scale=0
  $ 792 "Thread_1"
  thread Thread_1():
    while (True):
      $ 793 "If Start_thread≟ True "
      if (Start_thread ==   True  ):
        $ 794 "weight_value≔get_weight()"
        global weight_value=get_weight()
        $ 795 "diff≔target_weight-weight_value"
        global diff=target_weight-weight_value
        $ 796 "Wait: 0.2"
        sleep(0.2)
        $ 797 "sync()"
        sync()
      end
      $ 798 "sync()"
      sync()
    end
  end
  threadId_Thread_1 = run Thread_1()
  $ 799 "Thread_2"
  thread Thread_2():
    while (True):
      $ 800 "Loop vib_thread≟ True "
      thread Thread_while_800():
        while (True):
          $ 801 "diff≔target_weight-weight_value"
          global diff=target_weight-weight_value
          $ 802 "If diff>0.02 and spatula≠'spatula_flat_S'"
          global thread_flag_802=0
          thread Thread_if_802():
            $ 803 "vibration_4()"
            vibration_4()
            thread_flag_802 = 1
          end
          if (diff>0.02  and  spatula != "spatula_flat_S"):
            global thread_handler_802=run Thread_if_802()
            while (thread_flag_802 == 0):
              if not(diff>0.02  and  spatula != "spatula_flat_S"):
                kill thread_handler_802
                thread_flag_802 = 2
              else:
                sync()
              end
            end
          else:
            thread_flag_802 = 2
          end
          if (thread_flag_802 == 2):
            $ 805 "ElseIf diff>0.02 and spatula≟'spatula_flat_S'"
            if (diff>0.02 and spatula == "spatula_flat_S"):
              $ 806 "vibration_3()"
              vibration_3()
            else:
              $ 807 "ElseIf diff≤0.03"
              global thread_flag_807=0
              thread Thread_if_807():
                $ 808 "vibration_2()"
                vibration_2()
                thread_flag_807 = 1
              end
              if (diff <= 0.03):
                global thread_handler_807=run Thread_if_807()
                while (thread_flag_807 == 0):
                  if not(diff <= 0.03):
                    kill thread_handler_807
                    thread_flag_807 = 2
                  else:
                    sync()
                  end
                end
              else:
                thread_flag_807 = 2
              end
              if (thread_flag_807 == 2):
                $ 809 "Else" "noBreak"
                $ 810 "Set AO[0]=0.0"
                set_standard_analog_out(0, 0.0)
              end
            end
          end
        end
      end
      if (vib_thread ==   True  ):
        global thread_handler_800=run Thread_while_800()
        while (vib_thread ==   True  ):
          sync()
        end
        kill thread_handler_800
      end
      $ 811 "sync()"
      sync()
    end
  end
  threadId_Thread_2 = run Thread_2()
  while (True):
    $ 101 "Robot Program"
    $ 102 "MAIN"
    $ 103 "command_manager(external_control='uGO', cond_suspend=(ITM_Manipulated and AMR_AtTarget and AMR_Charging and AMR_Battery<40), cond_unsuspend=(AMR_Battery≟60))"
    command_manager(external_control="uGO", cond_suspend=(ITM_Manipulated  and  AMR_AtTarget  and  AMR_Charging  and  AMR_Battery<40), cond_unsuspend=(AMR_Battery == 60))
    $ 104 "log_state(STATE_Info)"
    log_state(STATE_Info)
    $ 105 "Switch STATE"
    switch_1 = STATE
    $ 106 "Case 1"
    if (1 == switch_1):
      $ 107 "Stopping"
      $ 108 "STATE_Info≔'Stopping'"
      global STATE_Info="Stopping"
      $ 109 "end_freedrive_mode()"
      end_freedrive_mode()
      $ 110 "Set"
      set_tcp(p[0.0,0.0,0.161,3.1415,0.0,0.0])
      $ 111 "PSE_T≔get_tool_free_pose(dir=[0,0,0.150], move_in_base_frame=True)"
      global PSE_T=get_tool_free_pose(dir=[0,0,0.150], move_in_base_frame=True)
      $ 112 "If is_reachable(Base_const, [PSE_T])"
      if (is_reachable(p[0.0,0.0,0.0,0.0,0.0,0.0], [PSE_T])):
        $ 113 "MoveL"
        $ 114 "PSE_T" "breakAfter"
        movel(PSE_T, a=1.2, v=0.15)
      end
      $ 115 "do_transition(keep_rxry=OBJ_Picked, r=0)"
      do_transition(keep_rxry=OBJ_Picked, r=0)
      $ 124 "Call Sub_AMR_MiR_V3"
      Sub_AMR_MiR_V3()
      $ 125 "If stopping() and AMR_Done"
      if (stopping()  and  AMR_Done):
        $ 126 "STATE≔2"
        global STATE=2
        $ 127 "ugo_update_outputs()"
        ugo_update_outputs()
      end
    elif (2 == switch_1):
      $ 128 "Case 2"
      $ 129 "Stopped"
      $ 130 "STATE_Info≔'Stopped'"
      global STATE_Info="Stopped"
      $ 131 "Call Sub_AMR_MiR_V3"
      Sub_AMR_MiR_V3()
      $ 132 "If CMD_Reset  or PB_Start"
      if (CMD_Reset   or  get_standard_digital_in(0)):
        $ 133 "STATE≔3"
        global STATE=3
        $ 134 "ugo_update_outputs()"
        ugo_update_outputs()
      end
    elif (3 == switch_1):
      $ 135 "Case 3"
      $ 136 " Resetting"
      $ 137 "STATE_Info≔'Resetting'"
      global STATE_Info="Resetting"
      $ 138 "uML"
      $ 139 "reset_error()"
      reset_error()
      $ 140 "reset_warning()"
      reset_warning()
      $ 141 "PROCESS_Step≔0"
      global PROCESS_Step=0
      $ 142 "PROCESS_Info≔''"
      global PROCESS_Info=""
      $ 143 "ARM_Referenced≔ False "
      global ARM_Referenced=  False
      $ 144 "WRK_Done≔ False "
      global WRK_Done=  False
      $ 145 "ITM_Prepared≔ False "
      global ITM_Prepared=  False
      $ 146 "ITM_Manipulated≔ False "
      global ITM_Manipulated=  False
      $ 147 "STP≔0"
      global STP=0
      $ 148 "Action≔0"
      global Action=0
      $ 149 "Action_Info≔''"
      global Action_Info=""
      $ 150 "ITM_ID≔0"
      global ITM_ID=0
      $ 151 "JIG≔0"
      global JIG=0
      $ 152 "JIG_Slot≔0"
      global JIG_Slot=0
      $ 153 "Task_info≔''"
      global Task_info=""
      $ 154 "Set"
      set_tcp(p[0.0,0.0,0.161,3.1415,0.0,0.0])
      $ 155 "App"
      $ 156 "'ADD APPLICATION SPECIFIC COMMANDS'"
      # 'ADD APPLICATION SPECIFIC COMMANDS'
      $ 157 "OBJ_Type≔0"
      global OBJ_Type=0
      $ 158 "OBJ_Nbr≔0"
      global OBJ_Nbr=0
      $ 159 "If CNT_Rack_Output≥50"
      if (CNT_Rack_Output >= 50):
        $ 160 "CNT_Rack_Output≔0"
        global CNT_Rack_Output=0
      end
      $ 161 "TASK≔struct(ID=0, NAVI=struct(target=0, footprint=0, protectiveOff=0, dock=0), WORK=struct(ITM_ID_Src=0, JIG_ID_Src=0, OBJ_Nbr_Src=0, ACT_Src=0, ITM_ID_Tgt=0, JIG_ID_Tgt=0, OBJ_Nbr_Tgt=0, ACT_Tgt=0, OBJ_Type=0))"
      global TASK=struct(ID=0, NAVI=struct(target=0, footprint=0, protectiveOff=0, dock=0), WORK=struct(ITM_ID_Src=0, JIG_ID_Src=0, OBJ_Nbr_Src=0, ACT_Src=0, ITM_ID_Tgt=0, JIG_ID_Tgt=0, OBJ_Nbr_Tgt=0, ACT_Tgt=0, OBJ_Type=0))
      $ 162 "Call Sub_AMR_MiR_V3"
      Sub_AMR_MiR_V3()
      $ 163 "If resetting() and AMR_Done"
      if (resetting()  and  AMR_Done):
        $ 164 "STATE≔4"
        global STATE=4
        $ 165 "ugo_update_outputs()"
        ugo_update_outputs()
      end
    elif (4 == switch_1):
      $ 166 "Case 4"
      $ 167 "Idle"
      $ 168 "STATE_Info≔'Idle'"
      global STATE_Info="Idle"
      $ 169 "If CMD_Start"
      if (CMD_Start):
        $ 170 "STATE≔5"
        global STATE=5
        $ 171 "ugo_update_outputs()"
        ugo_update_outputs()
      end
    elif (5 == switch_1):
      $ 172 "Case 5"
      $ 173 "Starting"
      $ 174 "STATE_Info≔'Starting'"
      global STATE_Info="Starting"
      $ 175 "'ADD COMMANDS WHAT TO START WITH'"
      # 'ADD COMMANDS WHAT TO START WITH'
      $ 176 "Call Sub_AMR_MiR_V3"
      Sub_AMR_MiR_V3()
      $ 177 "get ugo data"
      $ 178 "Assign Tasks"
      $ 179 "TASK.ID = ugo_get_task()"
      TASK.ID = ugo_get_task()
      $ 180 "If TASK.ID≟1"
      if (TASK.ID == 1):
        $ 181 "Task_info≔'Charge'"
        global Task_info="Charge"
        $ 182 "Parameters"
        $ 183 "AMR_PosTarget≔1"
        global AMR_PosTarget=1
      else:
        $ 184 "ElseIf TASK.ID≟9"
        if (TASK.ID == 9):
          $ 185 "'Pick Sarstedt Rack from Variable source'"
          # 'Pick Sarstedt Rack from Variable source'
          $ 186 "Task_info≔'Navigate to Target'"
          global Task_info="Navigate to Target"
          $ 187 "Parameters"
          $ 188 "AMR_PosTarget≔UGO.read_input('00','ITM_ID')"
          global AMR_PosTarget=UGO.read_input("00","ITM_ID")
        else:
          $ 189 "ElseIf TASK.ID≟13"
          if (TASK.ID == 13):
            $ 190 "Task_info≔'Dose Powder'"
            global Task_info="Dose Powder"
            $ 191 "Parameters"
            $ 192 "ITM_ID≔1"
            global ITM_ID=1
            $ 193 "W_now≔(UGO.read_input('00','Container_weight'))/1000"
            global W_now=(UGO.read_input("00","Container_weight"))/1000
            $ 194 "Pow_name≔(UGO.read_input('00','Powder_name'))"
            global Pow_name=(UGO.read_input("00","Powder_name"))
            $ 195 "target_weight≔(UGO.read_input('00','Target_weight'))/1000"
            global target_weight=(UGO.read_input("00","Target_weight"))/1000
            $ 196 "send_picking_info(Pow_name,target_weight)"
            send_picking_info(Pow_name,target_weight)
            $ 197 "OBJ_Type≔6"
            global OBJ_Type=6
            $ 198 "JIG≔17"
            global JIG=17
            $ 199 "AMR_PosTarget≔5"
            global AMR_PosTarget=5
          else:
            $ 200 "ElseIf TASK.ID≟49"
            if (TASK.ID == 49):
              $ 201 "Task_info≔'Pick Containers'"
              global Task_info="Pick Containers"
              $ 202 "Parameters"
              $ 203 "ITM_ID≔1"
              global ITM_ID=1
              $ 204 "OBJ_Type≔6"
              global OBJ_Type=6
              $ 205 "JIG≔15"
              global JIG=15
              $ 206 "AMR_PosTarget≔3"
              global AMR_PosTarget=3
            else:
              $ 207 "ElseIf TASK.ID≟50"
              if (TASK.ID == 50):
                $ 208 "Task_info≔'Decap Containers'"
                global Task_info="Decap Containers"
                $ 209 "Parameters"
                $ 210 "ITM_ID≔1"
                global ITM_ID=1
                $ 211 "OBJ_Type≔6"
                global OBJ_Type=6
                $ 212 "JIG≔16"
                global JIG=16
                $ 213 "AMR_PosTarget≔5"
                global AMR_PosTarget=5
              else:
                $ 214 "ElseIf TASK.ID≟51"
                if (TASK.ID == 51):
                  $ 215 "Task_info≔'Detect Spatula and transfer powder'"
                  global Task_info="Detect Spatula and transfer powder"
                  $ 216 "Parameters"
                  $ 217 "ITM_ID≔1"
                  global ITM_ID=1
                  $ 218 "target_weight≔(UGO.read_input('00','Target_weight'))/1000"
                  global target_weight=(UGO.read_input("00","Target_weight"))/1000
                  $ 219 "OBJ_Type≔8"
                  global OBJ_Type=8
                  $ 220 "JIG≔16"
                  global JIG=16
                  $ 221 "AMR_PosTarget≔5"
                  global AMR_PosTarget=5
                else:
                  $ 222 "ElseIf TASK.ID≟52"
                  if (TASK.ID == 52):
                    $ 223 "Task_info≔'Pick Powder'"
                    global Task_info="Pick Powder"
                    $ 224 "Parameters"
                    $ 225 "ITM_ID≔1"
                    global ITM_ID=1
                    $ 227 "OBJ_Type≔6"
                    global OBJ_Type=6
                    $ 228 "JIG≔15"
                    global JIG=15
                    $ 229 "AMR_PosTarget≔3"
                    global AMR_PosTarget=3
                  else:
                    $ 230 "ElseIf TASK.ID≟53"
                    if (TASK.ID == 53):
                      $ 231 "Task_info≔'Decap Powder'"
                      global Task_info="Decap Powder"
                      $ 232 "Parameters"
                      $ 233 "ITM_ID≔1"
                      global ITM_ID=1
                      $ 234 "OBJ_Type≔6"
                      global OBJ_Type=6
                      $ 235 "JIG≔1"
                      global JIG=1
                      $ 236 "AMR_PosTarget≔5"
                      global AMR_PosTarget=5
                    else:
                      $ 237 "ElseIf TASK.ID≟54"
                      if (TASK.ID == 54):
                        $ 238 "Task_info≔'Empty and swap Powder container'"
                        global Task_info="Empty and swap Powder container"
                        $ 247 "Parameters"
                        $ 248 "ITM_ID≔1"
                        global ITM_ID=1
                        $ 250 "W_now≔(UGO.read_input('00','Container_weight'))/1000"
                        global W_now=(UGO.read_input("00","Container_weight"))/1000
                        $ 251 "Pow_name≔(UGO.read_input('00','Powder_name'))"
                        global Pow_name=(UGO.read_input("00","Powder_name"))
                        $ 254 "OBJ_Type≔6"
                        global OBJ_Type=6
                        $ 255 "JIG≔17"
                        global JIG=17
                        $ 256 "AMR_PosTarget≔5"
                        global AMR_PosTarget=5
                      else:
                        $ 257 "ElseIf TASK.ID≟55"
                        if (TASK.ID == 55):
                          $ 258 "Task_info≔'Place Powder'"
                          global Task_info="Place Powder"
                          $ 259 "Parameters"
                          $ 260 "ITM_ID≔1"
                          global ITM_ID=1
                          $ 261 "OBJ_Type≔6"
                          global OBJ_Type=6
                          $ 262 "JIG≔21"
                          global JIG=21
                          $ 263 "AMR_PosTarget≔5"
                          global AMR_PosTarget=5
                        else:
                          $ 264 "ElseIf TASK.ID≟56"
                          if (TASK.ID == 56):
                            $ 265 "Task_info≔'Dose Powder'"
                            global Task_info="Dose Powder"
                            $ 266 "Parameters"
                            $ 267 "ITM_ID≔1"
                            global ITM_ID=1
                            $ 268 "target_weight≔(UGO.read_input('00','Target_weight'))/1000"
                            global target_weight=(UGO.read_input("00","Target_weight"))/1000
                            $ 269 "W_now≔(UGO.read_input('00','Container_weight'))/1000"
                            global W_now=(UGO.read_input("00","Container_weight"))/1000
                            $ 270 "Pow_name≔(UGO.read_input('00','Powder_name'))"
                            global Pow_name=(UGO.read_input("00","Powder_name"))
                            $ 271 "OBJ_Type≔6"
                            global OBJ_Type=6
                            $ 272 "JIG≔17"
                            global JIG=17
                            $ 273 "AMR_PosTarget≔5"
                            global AMR_PosTarget=5
                          else:
                            $ 274 "ElseIf TASK.ID≟57"
                            if (TASK.ID == 57):
                              $ 275 "Task_info≔'Recipe Powder dosing'"
                              global Task_info="Recipe Powder dosing"
                              $ 276 "Parameters"
                              $ 277 "ITM_ID≔1"
                              global ITM_ID=1
                              $ 278 "Pow_A≔(UGO.read_input('00','PowderA'))"
                              global Pow_A=(UGO.read_input("00","PowderA"))
                              $ 279 "Pow_B≔(UGO.read_input('00','PowderB'))"
                              global Pow_B=(UGO.read_input("00","PowderB"))
                              $ 280 "Pow_C≔(UGO.read_input('00','PowderC'))"
                              global Pow_C=(UGO.read_input("00","PowderC"))
                              $ 281 "Total_weight≔(UGO.read_input('00','Total_weight'))/1000"
                              global Total_weight=(UGO.read_input("00","Total_weight"))/1000
                              $ 282 "Pow_A_percent≔(UGO.read_input('00','PowderA_percentage'))/100"
                              global Pow_A_percent=(UGO.read_input("00","PowderA_percentage"))/100
                              $ 283 "Pow_B_percent≔(UGO.read_input('00','PowderB_percentage'))/100"
                              global Pow_B_percent=(UGO.read_input("00","PowderB_percentage"))/100
                              $ 284 "Pow_C_percent≔(UGO.read_input('00','PowderC_percentage'))/100"
                              global Pow_C_percent=(UGO.read_input("00","PowderC_percentage"))/100
                              $ 285 "OBJ_Type≔6"
                              global OBJ_Type=6
                              $ 286 "JIG≔17"
                              global JIG=17
                              $ 287 "AMR_PosTarget≔5"
                              global AMR_PosTarget=5
                            else:
                              $ 288 "ElseIf TASK.ID≟58"
                              if (TASK.ID == 58):
                                $ 289 "Task_info≔'Pick Powder containers'"
                                global Task_info="Pick Powder containers"
                                $ 290 "Parameters"
                                $ 291 "ITM_ID≔1"
                                global ITM_ID=1
                                $ 292 "OBJ_Type≔6"
                                global OBJ_Type=6
                                $ 293 "JIG≔15"
                                global JIG=15
                                $ 294 "AMR_PosTarget≔3"
                                global AMR_PosTarget=3
                              else:
                                $ 295 "Else" "noBreak"
                                $ 296 "set_error(ERROR_WRONG_ORDER)"
                                set_error(ERROR_WRONG_ORDER)
                              end
                            end
                          end
                        end
                      end
                    end
                  end
                end
              end
            end
          end
        end
      end
      $ 297 "test ugo"
      $ 298 "Wait: 0.2"
      sleep(0.2)
      $ 299 "ugo_update_outputs()"
      ugo_update_outputs()
      $ 300 "If starting() and AMR_Done"
      if (starting()  and  AMR_Done):
        $ 301 "log_message(Task_info, 'New Task: ')"
        log_message(Task_info, "New Task: ")
        $ 302 "log_message(to_str(TASK.ID), 'Task_ID: ')"
        log_message(to_str(TASK.ID), "Task_ID: ")
        $ 303 "do_transition(keep_rxry=OBJ_Picked)"
        do_transition(keep_rxry=OBJ_Picked)
        $ 304 "STATE≔6"
        global STATE=6
        $ 305 "ugo_update_outputs()"
        ugo_update_outputs()
      end
    elif (6 == switch_1):
      $ 306 "Case 6"
      $ 307 "Execute"
      $ 308 "STATE_Info≔'Execute'"
      global STATE_Info="Execute"
      $ 309 "If  not CMD_Hold and not CMD_Suspend"
      global thread_flag_309=0
      thread Thread_if_309():
        $ 310 "Switch PROCESS_Step"
        switch_2 = PROCESS_Step
        $ 311 "Case 0"
        if (0 == switch_2):
          $ 312 "PROCESS_Info≔'process control'"
          global PROCESS_Info="process control"
          $ 313 "log_process(PROCESS_Info)"
          log_process(PROCESS_Info)
          $ 314 "process control"
          $ 315 "If  not AMR_AtTarget"
          if (  not  AMR_AtTarget):
            $ 316 "PROCESS_Step≔1"
            global PROCESS_Step=1
          else:
            $ 317 "ElseIf (( not ITM_Prepared and  not WRK_Done) or (ITM_Prepared and WRK_Done))"
            if (((  not  ITM_Prepared  and    not  WRK_Done)  or  (ITM_Prepared  and  WRK_Done))):
              $ 318 "PROCESS_Step≔2"
              global PROCESS_Step=2
            else:
              $ 319 "ElseIf  not WRK_Done"
              if (  not  WRK_Done):
                $ 320 "PROCESS_Step≔3"
                global PROCESS_Step=3
              else:
                $ 321 "Else" "noBreak"
                $ 322 "task finished"
                $ 323 "PROCESS_Info≔''"
                global PROCESS_Info=""
                $ 324 "STATE≔7"
                global STATE=7
                $ 325 "ugo_update_outputs()"
                ugo_update_outputs()
              end
            end
          end
        elif (1 == switch_2):
          $ 326 "Case 1"
          $ 327 "navigate"
          $ 328 "'MOVING THE uML'"
          # 'MOVING THE uML'
          $ 329 "PROCESS_Info≔'move to target'"
          global PROCESS_Info="move to target"
          $ 330 "log_process(PROCESS_Info)"
          log_process(PROCESS_Info)
          $ 331 "If TASK.ID≟1"
          if (TASK.ID == 1):
            $ 332 "Action≔51"
            global Action=51
          else:
            $ 333 "Else" "noBreak"
            $ 334 "Action≔52"
            global Action=52
          end
          $ 335 "Call Sub_AMR_MiR_V3"
          Sub_AMR_MiR_V3()
          $ 336 "If AMR_Done"
          if (AMR_Done):
            $ 337 "PROCESS_Step≔0"
            global PROCESS_Step=0
          end
        elif (2 == switch_2):
          $ 338 "Case 2"
          $ 339 "prepare"
          $ 340 "'THINGS THAT HAVE TO BE DONE ONCE IN A SEQUENCE,WORKFLOW'"
          # 'THINGS THAT HAVE TO BE DONE ONCE IN A SEQUENCE,WORKFLOW'
          $ 341 "PROCESS_Info≔'prepare for work'"
          global PROCESS_Info="prepare for work"
          $ 342 "log_process(PROCESS_Info)"
          log_process(PROCESS_Info)
          $ 343 "If TASK.WORK.ITM_ID_Src>1"
          if (TASK.WORK.ITM_ID_Src>1):
            $ 344 "ITM_ID≔TASK.WORK.ITM_ID_Src"
            global ITM_ID=TASK.WORK.ITM_ID_Src
          else:
            $ 345 "ElseIf TASK.WORK.ITM_ID_Tgt>1"
            if (TASK.WORK.ITM_ID_Tgt>1):
              $ 346 "ITM_ID≔TASK.WORK.ITM_ID_Tgt"
              global ITM_ID=TASK.WORK.ITM_ID_Tgt
            end
          end
          $ 347 "If  not ARM_Referenced and (ITM_ID≠0)"
          if (  not  ARM_Referenced  and  (ITM_ID != 0)):
            $ 348 "STP≔1"
            global STP=1
          else:
            $ 349 "ElseIf ARM_Referenced or (ITM_ID≟0)"
            if (ARM_Referenced  or  (ITM_ID == 0)):
              $ 350 "STP≔2"
              global STP=2
            end
          end
          $ 351 "Switch STP"
          switch_3 = STP
          $ 352 "Case 1"
          if (1 == switch_3):
            $ 353 "reference"
            $ 354 "STP_Info≔'reference at target position'"
            global STP_Info="reference at target position"
            $ 355 "log_step(STP_Info)"
            log_step(STP_Info)
            $ 356 "If ITM_ID≟1"
            if (ITM_ID == 1):
              $ 357 "CAM_Done≔ True "
              global CAM_Done=  True
            else:
              $ 358 "Else" "noBreak"
              $ 359 "Action≔131"
              global Action=131
              $ 360 "Call Sub_Vision_V18"
              Sub_Vision_V18()
            end
            $ 362 "If CAM_Done and  not ERROR.FLAG"
            if (CAM_Done  and    not  ERROR.FLAG):
              $ 363 "log_step('ARM referenced')"
              log_step("ARM referenced")
              $ 364 "ARM_Referenced≔ True "
              global ARM_Referenced=  True
            end
          elif (2 == switch_3):
            $ 365 "Case 2"
            $ 366 "manipulate"
            $ 367 "STP_Info≔'manipulate item'"
            global STP_Info="manipulate item"
            $ 368 "log_step(STP_Info)"
            log_step(STP_Info)
            $ 369 "'In case pressing button is needed'"
            # 'In case pressing button is needed'
            $ 370 "If found_in_list(ITM_ID, ITM_ID_List)"
            if (found_in_list(ITM_ID, ITM_ID_List)):
              $ 371 "Switch ITM_ID"
              switch_4 = ITM_ID
              $ 372 "Case 0"
              if (0 == switch_4):
                $ 373 "ITM_Manipulated≔ not ITM_Manipulated"
                global ITM_Manipulated=  not  ITM_Manipulated
              elif (1 == switch_4):
                $ 374 "Case 1"
                $ 375 "ITM_Manipulated≔ not ITM_Manipulated"
                global ITM_Manipulated=  not  ITM_Manipulated
              elif (2 == switch_4):
                $ 376 "Case 2"
              else:
                $ 386 "Default Case"
                $ 387 "ITM_Manipulated≔ not ITM_Manipulated"
                global ITM_Manipulated=  not  ITM_Manipulated
              end
            end
          end
          $ 388 "ITM_Prepared≔(ITM_Manipulated or  not found_in_list(ITM_ID, ITM_ID_List)) and (ARM_Referenced or ITM_ID≟0) and  not WRK_Done"
          global ITM_Prepared=(ITM_Manipulated  or    not  found_in_list(ITM_ID, ITM_ID_List))  and  (ARM_Referenced  or  ITM_ID == 0)  and    not  WRK_Done
          $ 389 "STP≔0"
          global STP=0
          $ 390 "STP_Info≔''"
          global STP_Info=""
          $ 391 "PROCESS_Step≔0"
          global PROCESS_Step=0
        elif (3 == switch_2):
          $ 392 "Case 3"
          $ 393 "work"
          $ 394 "'ADD EVERY MACHINE, OBJECT, STATION TO WORK ON'"
          # 'ADD EVERY MACHINE, OBJECT, STATION TO WORK ON'
          $ 395 "Switch ITM_ID"
          switch_3 = ITM_ID
          $ 396 "Case 1"
          if (1 == switch_3):
            $ 397 "uLM"
            $ 398 "If TASK.ID≟12"
            if (TASK.ID == 12):
              $ 399 "fill racks"
              $ 400 "Action≔151"
              global Action=151
              $ 401 "Call Sub_Vision_V18"
              Sub_Vision_V18()
              $ 402 "If  not ERROR.FLAG"
              if (  not  ERROR.FLAG):
                $ 403 "Actions for the task"
                $ 404 "Action≔1"
                global Action=1
                $ 405 "JIG≔2"
                global JIG=2
                $ 406 "JIG_Slot≔CAM_Result[0]"
                global JIG_Slot=CAM_Result[0]
                $ 407 "OBJ_Nbr≔CAM_Result[0]"
                global OBJ_Nbr=CAM_Result[0]
                $ 408 "OBJ_Type≔2"
                global OBJ_Type=2
                $ 409 "Call Sub_Action_V4"
                Sub_Action_V4()
                $ 410 "If OBJ_Picked"
                if (OBJ_Picked):
                  $ 411 "CAM_Result.remove(0)"
                  CAM_Result.remove(0)
                  $ 412 "PRC_TubCounter≔PRC_TubCounter+1"
                  global PRC_TubCounter=PRC_TubCounter+1
                  $ 413 "If PRC_TubCounter%4≟0"
                  if (PRC_TubCounter%4 == 0):
                    $ 414 "JIG_Slot≔4"
                    global JIG_Slot=4
                  else:
                    $ 415 "Else" "noBreak"
                    $ 416 "JIG_Slot≔PRC_TubCounter%4"
                    global JIG_Slot=PRC_TubCounter%4
                  end
                  $ 417 "OBJ_Nbr≔ceil(PRC_TubCounter/4)"
                  global OBJ_Nbr=ceil(PRC_TubCounter/4)
                  $ 418 "Action≔2"
                  global Action=2
                  $ 419 "JIG≔4"
                  global JIG=4
                  $ 420 "Call Sub_Action_V4"
                  Sub_Action_V4()
                  $ 421 "Action≔151"
                  global Action=151
                  $ 422 "Call Sub_Vision_V18"
                  Sub_Vision_V18()
                end
              end
              $ 423 "If (CAM_Captures≥CAM_PRM_Retries) or (PRC_TubCounter≥32)"
              if ((CAM_Captures >= CAM_PRM_Retries)  or  (PRC_TubCounter >= 32)):
                $ 424 "PROCESS_Step≔0"
                global PROCESS_Step=0
                $ 425 "WRK_Done≔ True "
                global WRK_Done=  True
              end
            else:
              $ 426 "ElseIf TASK.ID≟13"
              if (TASK.ID == 13):
                $ 427 "Dose Powder"
                $ 428 "Action≔131"
                global Action=131
                $ 429 "Call Sub_Vision_V18"
                Sub_Vision_V18()
                $ 430 "Action≔34"
                global Action=34
                $ 431 "Call Sub_Action_V4"
                Sub_Action_V4()
                $ 432 "PROCESS_Step≔0"
                global PROCESS_Step=0
                $ 433 "WRK_Done≔ True "
                global WRK_Done=  True
              else:
                $ 434 "ElseIf TASK.ID≟49"
                if (TASK.ID == 49):
                  $ 435 "Pick Powder container"
                  $ 436 "Action≔131"
                  global Action=131
                  $ 437 "Call Sub_Vision_V18"
                  Sub_Vision_V18()
                  $ 438 "Action≔35"
                  global Action=35
                  $ 439 "Call Sub_Action_V4"
                  Sub_Action_V4()
                  $ 440 "PROCESS_Step≔0"
                  global PROCESS_Step=0
                  $ 441 "WRK_Done≔ True "
                  global WRK_Done=  True
                else:
                  $ 442 "ElseIf TASK.ID≟50"
                  if (TASK.ID == 50):
                    $ 443 "Decap containers"
                    $ 444 "Action≔36"
                    global Action=36
                    $ 445 "Call Sub_Action_V4"
                    Sub_Action_V4()
                    $ 446 "PROCESS_Step≔0"
                    global PROCESS_Step=0
                    $ 447 "WRK_Done≔ True "
                    global WRK_Done=  True
                  else:
                    $ 448 "ElseIf TASK.ID≟51"
                    if (TASK.ID == 51):
                      $ 449 "Detect Spatula and transfer powder"
                      $ 450 "Action≔131"
                      global Action=131
                      $ 451 "Call Sub_Vision_V18"
                      Sub_Vision_V18()
                      $ 452 "Action≔37"
                      global Action=37
                      $ 453 "Call Sub_Action_V4"
                      Sub_Action_V4()
                      $ 454 "PROCESS_Step≔0"
                      global PROCESS_Step=0
                      $ 455 "WRK_Done≔ True "
                      global WRK_Done=  True
                    else:
                      $ 456 "ElseIf TASK.ID≟52"
                      if (TASK.ID == 52):
                        $ 457 "Pick Powder container"
                        $ 458 "Action≔131"
                        global Action=131
                        $ 459 "Call Sub_Vision_V18"
                        Sub_Vision_V18()
                        $ 460 "Action≔39"
                        global Action=39
                        $ 461 "Call Sub_Action_V4"
                        Sub_Action_V4()
                        $ 462 "PROCESS_Step≔0"
                        global PROCESS_Step=0
                        $ 463 "WRK_Done≔ True "
                        global WRK_Done=  True
                      else:
                        $ 464 "ElseIf TASK.ID≟53"
                        if (TASK.ID == 53):
                          $ 465 "Decap containerA"
                          $ 466 "Action≔40"
                          global Action=40
                          $ 467 "Call Sub_Action_V4"
                          Sub_Action_V4()
                          $ 468 "PROCESS_Step≔0"
                          global PROCESS_Step=0
                          $ 469 "WRK_Done≔ True "
                          global WRK_Done=  True
                        else:
                          $ 470 "ElseIf TASK.ID≟55"
                          if (TASK.ID == 55):
                            $ 471 "Place Powder"
                            $ 472 "Action≔131"
                            global Action=131
                            $ 473 "Call Sub_Vision_V18"
                            Sub_Vision_V18()
                            $ 474 "Action≔41"
                            global Action=41
                            $ 475 "Call Sub_Action_V4"
                            Sub_Action_V4()
                            $ 476 "PROCESS_Step≔0"
                            global PROCESS_Step=0
                            $ 477 "WRK_Done≔ True "
                            global WRK_Done=  True
                          else:
                            $ 478 "ElseIf TASK.ID≟54"
                            if (TASK.ID == 54):
                              $ 479 "Empty and swap container"
                              $ 480 "Action≔131"
                              global Action=131
                              $ 481 "Call Sub_Vision_V18"
                              Sub_Vision_V18()
                              $ 482 "Action≔42"
                              global Action=42
                              $ 483 "Call Sub_Action_V4"
                              Sub_Action_V4()
                              $ 484 "PROCESS_Step≔0"
                              global PROCESS_Step=0
                              $ 485 "WRK_Done≔ True "
                              global WRK_Done=  True
                            else:
                              $ 486 "ElseIf TASK.ID≟56"
                              if (TASK.ID == 56):
                                $ 487 "Dispense Powder"
                                $ 488 "Action≔131"
                                global Action=131
                                $ 489 "Call Sub_Vision_V18"
                                Sub_Vision_V18()
                                $ 490 "Action≔43"
                                global Action=43
                                $ 491 "Call Sub_Action_V4"
                                Sub_Action_V4()
                                $ 492 "PROCESS_Step≔0"
                                global PROCESS_Step=0
                                $ 493 "WRK_Done≔ True "
                                global WRK_Done=  True
                              else:
                                $ 494 "ElseIf TASK.ID≟57"
                                if (TASK.ID == 57):
                                  $ 495 "Recipe Dosing"
                                  $ 496 "Action≔48"
                                  global Action=48
                                  $ 497 "Call Sub_Action_V4"
                                  Sub_Action_V4()
                                  $ 514 "PROCESS_Step≔0"
                                  global PROCESS_Step=0
                                  $ 515 "WRK_Done≔ True "
                                  global WRK_Done=  True
                                else:
                                  $ 516 "ElseIf TASK.ID≟58"
                                  if (TASK.ID == 58):
                                    $ 517 "Pick Powder containers"
                                    $ 518 "Num_cont_picked≔0"
                                    global Num_cont_picked=0
                                    $ 519 "powder_position≔'Position1'"
                                    global powder_position="Position1"
                                    $ 520 "Loop Num_cont_picked<3"
                                    while (Num_cont_picked<3):
                                      $ 521 "Action≔131"
                                      global Action=131
                                      $ 522 "Call Sub_Vision_V18"
                                      Sub_Vision_V18()
                                      $ 523 "Action≔47"
                                      global Action=47
                                      $ 524 "Call Sub_Action_V4"
                                      Sub_Action_V4()
                                    end
                                    $ 525 "PROCESS_Step≔0"
                                    global PROCESS_Step=0
                                    $ 526 "WRK_Done≔ True "
                                    global WRK_Done=  True
                                  end
                                end
                              end
                            end
                          end
                        end
                      end
                    end
                  end
                end
              end
            end
          elif (2 == switch_3):
            $ 527 "Case 2"
          elif (5 == switch_3):
            $ 569 "Case 5"
          elif (20 == switch_3):
            $ 577 "Case 20"
          elif (43 == switch_3):
            $ 639 "Case 43"
          else:
            $ 647 "Default Case"
            $ 648 "WRK_Done≔ True "
            global WRK_Done=  True
            $ 649 "PROCESS_Step≔0"
            global PROCESS_Step=0
          end
        end
        thread_flag_309 = 1
      end
      if (  not  CMD_Hold and not CMD_Suspend):
        global thread_handler_309=run Thread_if_309()
        while (thread_flag_309 == 0):
          if not(  not  CMD_Hold and not CMD_Suspend):
            kill thread_handler_309
            thread_flag_309 = 2
          else:
            sync()
          end
        end
      else:
        thread_flag_309 = 2
      end
      $ 650 "If CMD_Hold"
      if (CMD_Hold):
        $ 651 "STATE≔9"
        global STATE=9
        $ 652 "ugo_update_outputs()"
        ugo_update_outputs()
      else:
        $ 653 "ElseIf CMD_Suspend"
        if (CMD_Suspend):
          $ 654 "STATE≔12"
          global STATE=12
          $ 655 "ugo_update_outputs()"
          ugo_update_outputs()
        end
      end
    elif (7 == switch_1):
      $ 656 "Case 7"
      $ 657 "Completing"
      $ 658 "STATE_Info≔'Completing'"
      global STATE_Info="Completing"
      $ 659 "'ADD COMMANDS FOR COMPLETING THE PROCESS'"
      # 'ADD COMMANDS FOR COMPLETING THE PROCESS'
      $ 660 "do_transition(keep_rxry=OBJ_Picked)"
      do_transition(keep_rxry=OBJ_Picked)
      $ 661 "Call Sub_AMR_MiR_V3"
      Sub_AMR_MiR_V3()
      $ 662 "If completing() and AMR_Done"
      if (completing()  and  AMR_Done):
        $ 663 "STATE≔8"
        global STATE=8
        $ 664 "ugo_update_outputs()"
        ugo_update_outputs()
      end
    elif (8 == switch_1):
      $ 665 "Case 8"
      $ 666 "Complete"
      $ 667 "STATE_Info≔'Complete'"
      global STATE_Info="Complete"
      $ 668 "If CMD_Reset"
      if (CMD_Reset):
        $ 669 "STATE≔3"
        global STATE=3
        $ 670 "ugo_update_outputs()"
        ugo_update_outputs()
      end
    elif (9 == switch_1):
      $ 671 "Case 9"
      $ 672 "Holding"
      $ 673 "STATE_Info≔'Holding'"
      global STATE_Info="Holding"
      $ 674 "stopl(0.5)"
      stopl(0.5)
      $ 675 "Call Sub_AMR_MiR_V3"
      Sub_AMR_MiR_V3()
      $ 676 "If holding() and AMR_Done"
      if (holding()  and  AMR_Done):
        $ 677 "STATE≔10"
        global STATE=10
        $ 678 "ugo_update_outputs()"
        ugo_update_outputs()
      end
    elif (10 == switch_1):
      $ 679 "Case 10"
      $ 680 "Held"
      $ 681 "STATE_Info≔'Held'"
      global STATE_Info="Held"
      $ 682 "If CMD_Unhold"
      if (CMD_Unhold):
        $ 683 "end_freedrive_mode()"
        end_freedrive_mode()
        $ 684 "STATE≔11"
        global STATE=11
        $ 685 "ugo_update_outputs()"
        ugo_update_outputs()
      else:
        $ 686 "ElseIf FNC_Freedrive"
        if (FNC_Freedrive):
          $ 687 "freedrive_mode()"
          freedrive_mode()
        else:
          $ 688 "Else" "noBreak"
          $ 689 "end_freedrive_mode()"
          end_freedrive_mode()
        end
      end
    elif (11 == switch_1):
      $ 690 "Case 11"
      $ 691 "Unholding"
      $ 692 "STATE_Info≔'Unholding'"
      global STATE_Info="Unholding"
      $ 693 "Clearing"
      $ 694 "Switch ERROR.ID"
      switch_2 = ERROR.ID
      $ 695 "Case 1002"
      if (1002 == switch_2):
        $ 696 "AMR_AtTarget≔ False "
        global AMR_AtTarget=  False
        $ 697 "ARM_Referenced≔ False "
        global ARM_Referenced=  False
        $ 698 "ITM_Prepared≔ False "
        global ITM_Prepared=  False
        $ 699 "PROCESS_Step≔1"
        global PROCESS_Step=1
      elif (2007 == switch_2):
        $ 700 "Case 2007"
        $ 701 "PROCESS_Step≔1"
        global PROCESS_Step=1
      end
      $ 702 "reset_error()"
      reset_error()
      $ 703 "reset_warning()"
      reset_warning()
      $ 704 "OBJ_Picked≔gripper_has_object()"
      global OBJ_Picked=gripper_has_object()
      $ 705 "Call Sub_AMR_MiR_V3"
      Sub_AMR_MiR_V3()
      $ 706 "If unholding() and AMR_Done"
      if (unholding()  and  AMR_Done):
        $ 707 "STATE≔6"
        global STATE=6
        $ 708 "ugo_update_outputs()"
        ugo_update_outputs()
      end
    elif (12 == switch_1):
      $ 709 "Case 12"
      $ 710 "Suspending"
      $ 711 "STATE_Info≔'Suspending'"
      global STATE_Info="Suspending"
      $ 712 "PROCESS_Info≔str_cat(PROCESS_Info, ' suspended')"
      global PROCESS_Info=str_cat(PROCESS_Info, " suspended")
      $ 713 "If suspending()"
      if (suspending()):
        $ 714 "STATE≔13"
        global STATE=13
        $ 715 "ugo_update_outputs()"
        ugo_update_outputs()
      end
    elif (13 == switch_1):
      $ 716 "Case 13"
      $ 717 "Suspended"
      $ 718 "STATE_Info≔'Suspended'"
      global STATE_Info="Suspended"
      $ 719 "Call Sub_AMR_MiR_V3"
      Sub_AMR_MiR_V3()
      $ 720 "If CMD_Unsuspend"
      if (CMD_Unsuspend):
        $ 721 "STATE≔14"
        global STATE=14
        $ 722 "ugo_update_outputs()"
        ugo_update_outputs()
      end
    elif (14 == switch_1):
      $ 723 "Case 14"
      $ 724 "Unsuspending"
      $ 725 "STATE_Info≔'Unsuspending'"
      global STATE_Info="Unsuspending"
      $ 726 "PROCESS_Step≔0"
      global PROCESS_Step=0
      $ 727 "If unsuspending()"
      if (unsuspending()):
        $ 728 "STATE≔6"
        global STATE=6
        $ 729 "ugo_update_outputs()"
        ugo_update_outputs()
      end
    elif (15 == switch_1):
      $ 730 "Case 15"
      $ 731 "Aborting"
      $ 732 "STATE_Info≔'Aborting'"
      global STATE_Info="Aborting"
      $ 733 "If aborting()"
      if (aborting()):
        $ 734 "STATE≔16"
        global STATE=16
        $ 735 "ugo_update_outputs()"
        ugo_update_outputs()
      end
    elif (16 == switch_1):
      $ 736 "Case 16"
      $ 737 "Aborted"
      $ 738 "STATE_Info≔'Aborted'"
      global STATE_Info="Aborted"
      $ 739 "If CMD_Clear"
      if (CMD_Clear):
        $ 740 "STATE≔17"
        global STATE=17
        $ 741 "ugo_update_outputs()"
        ugo_update_outputs()
      end
    elif (17 == switch_1):
      $ 742 "Case 17"
      $ 743 "Clearing"
      $ 744 "STATE_Info≔'Clearing'"
      global STATE_Info="Clearing"
      $ 745 "Clearing"
      $ 746 "reset_warning()"
      reset_warning()
      $ 747 "reset_error()"
      reset_error()
      $ 748 "If clearing()"
      if (clearing()):
        $ 749 "STATE≔2"
        global STATE=2
        $ 750 "ugo_update_outputs()"
        ugo_update_outputs()
      end
    end
    $ 751 "log_state(STATE_Info)"
    log_state(STATE_Info)
    $ 752 "log_warning(WARNING.MSG)"
    log_warning(WARNING.MSG)
    $ 753 "log_error(ERROR.MSG)"
    log_error(ERROR.MSG)
    $ 754 "Times"
    $ 755 "Switch STATE"
    switch_1 = STATE
    $ 756 "Case 1"
    if (1 == switch_1):
      $ 757 "TM_St_Stopping≔get_time(STATE_Times[STATE-1])"
      global TM_St_Stopping=get_time(STATE_Times[STATE-1])
    elif (2 == switch_1):
      $ 758 "Case 2"
      $ 759 "TM_St_Stopped≔get_time(STATE_Times[STATE-1])"
      global TM_St_Stopped=get_time(STATE_Times[STATE-1])
    elif (3 == switch_1):
      $ 760 "Case 3"
      $ 761 "TM_St_Resetting≔get_time(STATE_Times[STATE-1])"
      global TM_St_Resetting=get_time(STATE_Times[STATE-1])
    elif (4 == switch_1):
      $ 762 "Case 4"
      $ 763 "TM_St_Idle≔get_time(STATE_Times[STATE-1])"
      global TM_St_Idle=get_time(STATE_Times[STATE-1])
    elif (5 == switch_1):
      $ 764 "Case 5"
      $ 765 "TM_St_Starting≔get_time(STATE_Times[STATE-1])"
      global TM_St_Starting=get_time(STATE_Times[STATE-1])
    elif (6 == switch_1):
      $ 766 "Case 6"
      $ 767 "TM_St_Execute≔get_time(STATE_Times[STATE-1])"
      global TM_St_Execute=get_time(STATE_Times[STATE-1])
    elif (7 == switch_1):
      $ 768 "Case 7"
      $ 769 "TM_St_Completin≔get_time(STATE_Times[STATE-1])"
      global TM_St_Completin=get_time(STATE_Times[STATE-1])
    elif (8 == switch_1):
      $ 770 "Case 8"
      $ 771 "TM_St_Complete≔get_time(STATE_Times[STATE-1])"
      global TM_St_Complete=get_time(STATE_Times[STATE-1])
    elif (9 == switch_1):
      $ 772 "Case 9"
      $ 773 "TM_St_Holding≔get_time(STATE_Times[STATE-1])"
      global TM_St_Holding=get_time(STATE_Times[STATE-1])
    elif (10 == switch_1):
      $ 774 "Case 10"
      $ 775 "TM_St_Held≔get_time(STATE_Times[STATE-1])"
      global TM_St_Held=get_time(STATE_Times[STATE-1])
    elif (11 == switch_1):
      $ 776 "Case 11"
      $ 777 "TM_St_Unholding≔get_time(STATE_Times[STATE-1])"
      global TM_St_Unholding=get_time(STATE_Times[STATE-1])
    elif (12 == switch_1):
      $ 778 "Case 12"
      $ 779 "TM_St_Suspendin≔get_time(STATE_Times[STATE-1])"
      global TM_St_Suspendin=get_time(STATE_Times[STATE-1])
    elif (13 == switch_1):
      $ 780 "Case 13"
      $ 781 "TM_St_Suspended≔get_time(STATE_Times[STATE-1])"
      global TM_St_Suspended=get_time(STATE_Times[STATE-1])
    elif (14 == switch_1):
      $ 782 "Case 14"
      $ 783 "TM_St_Unsuspend≔get_time(STATE_Times[STATE-1])"
      global TM_St_Unsuspend=get_time(STATE_Times[STATE-1])
    elif (15 == switch_1):
      $ 784 "Case 15"
      $ 785 "TM_St_Aborting≔get_time(STATE_Times[STATE-1])"
      global TM_St_Aborting=get_time(STATE_Times[STATE-1])
    elif (16 == switch_1):
      $ 786 "Case 16"
      $ 787 "TM_St_Aborted≔get_time(STATE_Times[STATE-1])"
      global TM_St_Aborted=get_time(STATE_Times[STATE-1])
    elif (17 == switch_1):
      $ 788 "Case 17"
      $ 789 "TM_St_Clearing≔get_time(STATE_Times[STATE-1])"
      global TM_St_Clearing=get_time(STATE_Times[STATE-1])
    end
    $ 791 "Wait: 0.1"
    sleep(0.1)
  end
end
